FUNCTION_BLOCK EQ_LinearAxis (* An equipment block: the only block that touches this equipment's pins. Skills send it what to switch over a local channel; it switches the outputs (off first, then on), reads the inputs every cycle and reports them to the skills and to OPC UA. One skill holds it at a time; on release or when the module aborts it switches everything off. Technical: Lift of the stoppering head, a stepper motor through a step and direction driver, with a limit switch at the top (home); equipment IO: owns its IO points, writes the output values its holder sends, reads its inputs every cycle and reports changes *)
  (* Standard: 61499-2 *)
  (* Version 0.1, 2026-09-28, Project contributors, AAU Smart Production Lab *)
  PACKAGE stoppering;
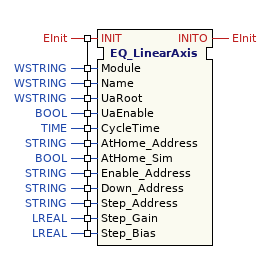
  EVENT_INPUT
    INIT : EInit WITH Module, Name, UaRoot, UaEnable, CycleTime, AtHome_Address, AtHome_Sim, Enable_Address, Down_Address, Step_Address, Step_Gain, Step_Bias; (* Initialise, once at start-up (the INIT chain); takes the values given with it *)
  END_EVENT
  EVENT_OUTPUT
    INITO : EInit; (* Initialised: the next block of the INIT chain goes on *)
  END_EVENT
  VAR_INPUT
    Module : WSTRING; (* The module's name; its local channels are named after it (loc[<Module>/...]) *)
    Name : WSTRING := "LinearAxis"; (* The equipment item's name: its local channels and OPC UA folder *)
    UaRoot : WSTRING; (* The module's OPC UA folder, e.g. /Objects/Filling *)
    UaEnable : BOOL; (* Publish on OPC UA *)
    CycleTime : TIME := T#50ms; (* How often the inputs are read *)
    AtHome_Address : STRING; (* Where AtHome is: 'gpio[chip:line(:pull_up|:pull_down)(:active_low)]', 'pwm[chip:channel:period_ns]', 'modbus[...]', 'sim', or an IO handle's name; empty: not connected *)
    AtHome_Sim : BOOL := FALSE; (* The value of AtHome when simulated (address 'sim') *)
    Enable_Address : STRING; (* Where Enable is: 'gpio[chip:line(:pull_up|:pull_down)(:active_low)]', 'pwm[chip:channel:period_ns]', 'modbus[...]', 'sim', or an IO handle's name; empty: not connected *)
    Down_Address : STRING; (* Where Down is: 'gpio[chip:line(:pull_up|:pull_down)(:active_low)]', 'pwm[chip:channel:period_ns]', 'modbus[...]', 'sim', or an IO handle's name; empty: not connected *)
    Step_Address : STRING; (* Where Step is: 'gpio[chip:line(:pull_up|:pull_down)(:active_low)]', 'pwm[chip:channel:period_ns]', 'modbus[...]', 'sim', or an IO handle's name; empty: not connected *)
    Step_Gain : LREAL := 655.35; (* Step: raw = Bias + value * Gain *)
    Step_Bias : LREAL := 0.0; (* Step: raw = Bias + value * Gain *)
  END_VAR
  (* Group Core: One holder at a time, break before make, all off on release or abort; scanned every CycleTime *)
  (* Group Channels: Local channels to and from the skills (cmd, release, state), the module's state, and the inputs over OPC UA *)
  (* Group Inputs: The equipment's sensors: read every cycle, one block per IO point *)
  (* Group Outputs: The equipment's actuators: written on a change and every cycle, one block per IO point *)
  FBS
    Logic : stoppering::EL_LinearAxis; (* The equipment's logic (EL_): takes commands from one holder at a time, switches the outputs (off first, then on), switches all off on release or module abort, and reports input changes. *) {SET_ATTRIBUTE(GroupName, Core)}
    Cycle : iec61499::events::E_CYCLE; (* Ticks every cycle so the inputs are read and the outputs refreshed. *) {SET_ATTRIBUTE(GroupName, Core)}
    MoveT : iec61499::events::E_DELAY; (* Times a move to a position: the distance divided by the axis' speed. *) {SET_ATTRIBUTE(GroupName, Core)}
    Mode : modlib::MOD_StateView; (* Watches the module's PackML state, to switch everything off when the module aborts. *) {SET_ATTRIBUTE(GroupName, Channels)}
    SubCmd : iec61499::net::SUBSCRIBE_8(QI := TRUE); (* Receives the commands skills send on this equipment's command channel. *) {SET_ATTRIBUTE(GroupName, Channels)}
    SubRelease : iec61499::net::SUBSCRIBE_1(QI := TRUE); (* Hears the module's release channel: when its holder gives up, everything goes off. *) {SET_ATTRIBUTE(GroupName, Channels)}
    PubState : iec61499::net::PUBLISH_5(QI := TRUE); (* Publishes the inputs and the holder on this equipment's state channel, for the skills. *) {SET_ATTRIBUTE(GroupName, Channels)}
    PubUa : iec61499::net::PUBLISH_4; (* Writes the inputs (and a position, if it keeps one) to OPC UA, below Equipment/<item>. *) {SET_ATTRIBUTE(GroupName, Channels)}
    In_AtHome : modlib::IO_DI; (* The pin AtHome: reads the input at AtHome_Address (a Pi pin, Modbus, or simulated). *) {SET_ATTRIBUTE(GroupName, Inputs)}
    Out_Enable : modlib::IO_DO; (* The pin Enable: switches the output at Enable_Address (a Pi pin, Modbus, or simulated). *) {SET_ATTRIBUTE(GroupName, Outputs)}
    Out_Down : modlib::IO_DO; (* The pin Down: switches the output at Down_Address (a Pi pin, Modbus, or simulated). *) {SET_ATTRIBUTE(GroupName, Outputs)}
    Out_Step : modlib::IO_AO; (* The pin Step: switches the output at Step_Address (a Pi pin, Modbus, or simulated). *) {SET_ATTRIBUTE(GroupName, Outputs)}
  END_FBS
  EVENT_CONNECTIONS
    Logic.MOVE_START TO MoveT.START;
    Logic.MOVE_STOP TO MoveT.STOP;
    MoveT.EO TO Logic.MOVE_T;
    INIT TO Logic.INIT;
    Logic.INITO TO Mode.INIT;
    Mode.INITO TO SubCmd.INIT;
    SubCmd.INITO TO SubRelease.INIT;
    SubRelease.INITO TO PubState.INIT;
    PubState.INITO TO PubUa.INIT;
    PubUa.INITO TO In_AtHome.INIT;
    In_AtHome.INITO TO Out_Enable.INIT;
    Out_Enable.INITO TO Out_Down.INIT;
    Out_Down.INITO TO Out_Step.INIT;
    Out_Step.INITO TO Cycle.START;
    Out_Step.INITO TO INITO;
    SubCmd.IND TO Logic.CMD;
    SubRelease.IND TO Logic.RELEASE;
    Mode.CHG TO Logic.MOD_CHG;
    Cycle.EO TO Logic.REFRESH;
    Cycle.EO TO In_AtHome.REQ;
    In_AtHome.CNF TO Logic.SAMPLE;
    Logic.STATE TO PubState.REQ;
    Logic.STATE TO PubUa.REQ;
    Logic.DRIVE TO Out_Enable.REQ;
    Out_Enable.CNF TO Out_Down.REQ;
    Out_Down.CNF TO Out_Step.REQ;
    Out_Step.CNF TO Logic.DRIVEN;
  END_CONNECTIONS
  DATA_CONNECTIONS
    Logic.MoveDT TO MoveT.DT;
    Module TO Logic.Module;
    Name TO Logic.Name;
    UaRoot TO Logic.UaRoot;
    Module TO Mode.Module;
    Logic.IdCmd TO SubCmd.ID;
    Logic.IdRelease TO SubRelease.ID;
    Logic.IdState TO PubState.ID;
    Logic.IdPub TO PubUa.ID;
    UaEnable TO PubUa.QI;
    CycleTime TO Cycle.DT;
    SubCmd.RD_1 TO Logic.C_Holder;
    SubCmd.RD_2 TO Logic.C_Release;
    SubCmd.RD_3 TO Logic.C_Enable;
    SubCmd.RD_4 TO Logic.C_Down;
    SubCmd.RD_5 TO Logic.C_Step;
    SubCmd.RD_6 TO Logic.CE_Step;
    SubCmd.RD_7 TO Logic.C_Move;
    SubCmd.RD_8 TO Logic.C_Goal;
    SubRelease.RD_1 TO Logic.R_Holder;
    Mode.State TO Logic.ModuleState;
    AtHome_Address TO In_AtHome.Address;
    AtHome_Sim TO In_AtHome.SimValue;
    In_AtHome.IN TO Logic.I_AtHome;
    Logic.AtHome TO PubState.SD_1;
    Logic.AtHome TO PubUa.SD_1;
    Logic.ActualPosition TO PubState.SD_2;
    Logic.ActualPosition TO PubUa.SD_2;
    Logic.Homed TO PubState.SD_3;
    Logic.Homed TO PubUa.SD_3;
    Logic.Moving TO PubState.SD_4;
    Logic.Moving TO PubUa.SD_4;
    Logic.Holder TO PubState.SD_5;
    Enable_Address TO Out_Enable.Address;
    Logic.O_Enable TO Out_Enable.OUT;
    Down_Address TO Out_Down.Address;
    Logic.O_Down TO Out_Down.OUT;
    Step_Address TO Out_Step.Address;
    Logic.O_Step TO Out_Step.OUT;
    Logic.E_Step TO Out_Step.EN;
    Step_Gain TO Out_Step.Gain;
    Step_Bias TO Out_Step.Bias;
  END_CONNECTIONS
END_FUNCTION_BLOCK
